Staubli VAL3: exercice4.pgx

program exercice4()
  local num l_nNbKapla
  local pointRx dest
  local trsf Pas
  local trsf Decal
begin
  Pas.x = (((Prise5[4].trsf.x)-(Prise5[0].trsf.x))/4)
  Pas.y = (((Prise5[4].trsf.y)-(Prise5[0].trsf.y))/4)
  Pas.z = (((Prise5[4].trsf.z)-(Prise5[0].trsf.z))/4)

  for l_nNbKapla = 0 to 4

    Decal.x = l_nNbKapla * Pas.x
    Decal.y = l_nNbKapla * Pas.y
    Decal.z = l_nNbKapla * Pas.z

    dest = compose(Prise5[0],world,Decal)

    movej(appro(dest,{0,0,-50,0,0,0}),tPince,mRapide)
    movel(dest,tPince,mLent)
    call fermerPince()
    movel(appro(dest,{0,0,-50,0,0,0}),tPince,mRapide)

    movej(jDepart,tPince,mRapide)
    movej(appro(pDepose[0],{0,0,-50,0,0,0}),tPince,mRapide)
    movel(pDepose[0],tPince,mLent)
    call ouvrirPince()
    movel(appro(pDepose,{0,0,-50,0,0,0}),tPince,mRapide)
    movej(jDepart,tPince,mLent)
    waitEndMove()
    delay(3)
    endFor

end
